// TIA Portal V21 export
FUNCTION "FC_AnaDead" : Int   // FC15, SCL
TITLE = Analyzer: dead block
{ S7_Optimized_Access := 'TRUE' }
// Rule C26k: no OB calls this block
// stored: SetENOAutomatically false
   VAR_INPUT
      Value : Int;   // Value
   END_VAR
BEGIN

       #FC_AnaDead := #Value + 1;
END_FUNCTION
